FUNCTION_BLOCK FB_LightCatalogTests EXTENDS TcUnit.FB_TestSuite
VAR
END_VAR

CatalogIsStableAndTracksLightOutputs();

METHOD PRIVATE CatalogIsStableAndTracksLightOutputs
VAR
    fbHome : FB_Home;
    stInputs : ST_HomeInputs;
    stOutputs : ST_HomeOutputs;
    nIndex : DINT;
    nOtherIndex : DINT;
    nFirstIndex : DINT;
    nLastIndex : DINT;
    nLightCount : DINT;
END_VAR
TEST('Light catalog identities are unique and snapshots track light outputs');

nFirstIndex := 1;
stInputs.Workshop.bButton := TRUE;
stInputs.Entryway.bLowerButton := TRUE;
stInputs.Entryway.bUpperButton := TRUE;
fbHome(stInputs := stInputs, stOutputs => stOutputs);
nLightCount := fbHome.nLightCount;
nLastIndex := nFirstIndex + nLightCount - 1;
AssertTrue(Condition := fbHome.nLightCount = (UPPER_BOUND(fbHome.aLights, 1) - LOWER_BOUND(fbHome.aLights, 1) + 1), Message := 'Reported catalog count matches the light array bounds');

FOR nIndex := nFirstIndex TO nLastIndex DO
    AssertTrue(Condition := fbHome.aLights[nIndex].sLocationId <> '', Message := 'Catalog location id is not empty');
    AssertTrue(Condition := fbHome.aLights[nIndex].sId <> '', Message := 'Catalog light id is not empty');
    AssertTrue(Condition := fbHome.aLights[nIndex].sType = 'light', Message := 'Catalog type is light');
    AssertFalse(Condition := fbHome.aLights[nIndex].bOn, Message := 'Startup-high input leaves catalog state off');
    FOR nOtherIndex := nIndex + 1 TO nLastIndex DO
        AssertFalse(Condition := fbHome.aLights[nIndex].sLocationId = fbHome.aLights[nOtherIndex].sLocationId AND fbHome.aLights[nIndex].sId = fbHome.aLights[nOtherIndex].sId, Message := 'Catalog location/id pairs are unique');
    END_FOR
END_FOR
AssertTrue(Condition := fbHome.aLights[1].sLocationId = 'H.01-09' AND fbHome.aLights[1].sId = 'main', Message := 'Workshop identity is configured');
AssertTrue(Condition := fbHome.aLights[2].sLocationId = 'H.01-01' AND fbHome.aLights[2].sId = 'main', Message := 'Entryway identity is configured');
AssertTrue(Condition := fbHome.aLights[3].sLocationId = 'H.01-01' AND fbHome.aLights[3].sId = 'temporary', Message := 'Temporary identity is configured');
AssertTrue(Condition := fbHome.nLightCount = 6 AND fbHome.bCatalogReady, Message := 'Catalog reports six ready lights');
AssertTrue(Condition := fbHome.aLights[4].sLocationId = 'H.01-02' AND fbHome.aLights[4].sId = 'main', Message := 'Hall group identity is configured');
AssertTrue(Condition := fbHome.aLights[5].sLocationId = 'H.01-02' AND fbHome.aLights[5].sId = 'outer_spots', Message := 'Hall outer spots identity is configured');
AssertTrue(Condition := fbHome.aLights[6].sLocationId = 'H.01-02' AND fbHome.aLights[6].sId = 'middle_spot', Message := 'Hall middle spot identity is configured');

stInputs.Workshop.bButton := FALSE;
stInputs.Entryway.bLowerButton := FALSE;
stInputs.Entryway.bUpperButton := FALSE;
fbHome(stInputs := stInputs, stOutputs => stOutputs);
stInputs.Workshop.bButton := TRUE;
stInputs.Entryway.bLowerButton := TRUE;
stInputs.Entryway.bUpperButton := TRUE;
fbHome(stInputs := stInputs, stOutputs => stOutputs);
AssertTrue(Condition := fbHome.aLights[1].bOn = stOutputs.Workshop.bLightRelay, Message := 'Workshop snapshot matches output in same scan');
AssertTrue(Condition := fbHome.aLights[2].bOn = stOutputs.Entryway.bLightRelay, Message := 'Entryway snapshot matches output in same scan');
AssertTrue(Condition := fbHome.aLights[3].bOn = stOutputs.Entryway.bTemporaryLightRelay, Message := 'Temporary snapshot matches output in same scan');
AssertTrue(Condition := fbHome.aLights[4].bOn = (stOutputs.Hall.bOuterSpotsRelay OR stOutputs.Hall.bMiddleSpotRelay), Message := 'Hall group snapshot is derived from members');
AssertTrue(Condition := fbHome.aLights[5].bOn = stOutputs.Hall.bOuterSpotsRelay, Message := 'Hall outer spots snapshot matches relay');
AssertTrue(Condition := fbHome.aLights[6].bOn = stOutputs.Hall.bMiddleSpotRelay, Message := 'Hall middle spot snapshot matches relay');
AssertTrue(Condition := fbHome.aLights[1].bOn AND fbHome.aLights[2].bOn AND fbHome.aLights[3].bOn, Message := 'Workshop and Entryway presses turn their lights on');
AssertTrue(Condition := fbHome.aLights[1].sLocationId = 'H.01-09' AND fbHome.aLights[1].sId = 'main', Message := 'Workshop identity survives toggle');
AssertTrue(Condition := fbHome.aLights[2].sLocationId = 'H.01-01' AND fbHome.aLights[2].sId = 'main', Message := 'Entryway identity survives toggle');
AssertTrue(Condition := fbHome.aLights[3].sLocationId = 'H.01-01' AND fbHome.aLights[3].sId = 'temporary', Message := 'Temporary identity survives toggle');
AssertTrue(Condition := fbHome.aLights[4].sLocationId = 'H.01-02' AND fbHome.aLights[4].sId = 'main', Message := 'Hall group identity survives toggle');
fbHome(stInputs := stInputs, stOutputs => stOutputs);
AssertTrue(Condition := fbHome.aLights[1].bOn AND fbHome.aLights[2].bOn AND fbHome.aLights[3].bOn, Message := 'Held Workshop and Entryway buttons do not toggle again');

stInputs.Workshop.bButton := FALSE;
stInputs.Entryway.bLowerButton := FALSE;
stInputs.Entryway.bUpperButton := FALSE;
fbHome(stInputs := stInputs, stOutputs => stOutputs);
stInputs.Workshop.bButton := TRUE;
stInputs.Entryway.bLowerButton := TRUE;
stInputs.Entryway.bUpperButton := TRUE;
fbHome(stInputs := stInputs, stOutputs => stOutputs);
AssertTrue(Condition := NOT fbHome.aLights[1].bOn AND NOT fbHome.aLights[2].bOn AND NOT fbHome.aLights[3].bOn, Message := 'Second Workshop and Entryway presses toggle their lights off');
AssertTrue(Condition := fbHome.aLights[1].bOn = stOutputs.Workshop.bLightRelay, Message := 'Workshop OFF snapshot matches output in same scan');
AssertTrue(Condition := fbHome.aLights[2].bOn = stOutputs.Entryway.bLightRelay, Message := 'Entryway OFF snapshot matches output in same scan');
AssertTrue(Condition := fbHome.aLights[3].bOn = stOutputs.Entryway.bTemporaryLightRelay, Message := 'Temporary OFF snapshot matches output in same scan');
AssertTrue(Condition := NOT fbHome.aLights[4].bOn AND NOT fbHome.aLights[5].bOn AND NOT fbHome.aLights[6].bOn, Message := 'Hall catalog remains off until Hall upper is pressed');

TEST_FINISHED();
END_METHOD

END_FUNCTION_BLOCK

(* stored: Version 1.1.0.1
   POU FB_LightCatalogTests: Id {08fdb221-4340-488f-bad9-a16217798d11}, SpecialFunc None
   Method CatalogIsStableAndTracksLightOutputs: Id {3f542897-b53f-4eb0-a2bb-873f7a568e3c} *)
